Staubli VAL3: setPageMaxJntForce.pgx

public program setPageMaxJntForce()
  local num i
begin
  //页面修改扭矩库限值
  if sArmType=="4_Axis"
    for i=0 to 3
      forcedata:tArm4Force[sArmDetail].nMaxJnt4Force[i]=nMaxJntForce[i]
    endFor
  elseIf sArmType=="6_Axis"
    for i=0 to 5
      forcedata:tArm6Force[sArmDetail].nMaxJnt6Force[i]=nMaxJntForce[i]
    endFor
  endIf
  forcedata:libSave()
  delay(0.1)
end
